// TIA Portal V21 export
FUNCTION_BLOCK "ClassicFbd"   // FB11, FBD
TITLE = ClassicFbd
// Function block diagram on a classic CPU.
   VAR_INPUT
      enable : Bool;
   END_VAR
   VAR_OUTPUT
      running : Bool;
   END_VAR
   VAR
      latched : Bool;
   END_VAR
BEGIN

REGION Network 1: Latch
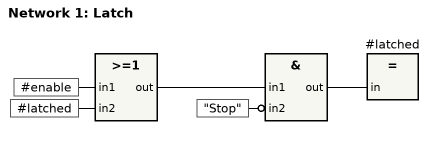
   #latched := (#enable OR #latched) AND NOT "Stop";
END_REGION
END_FUNCTION_BLOCK
